Fanuc KAREL source: KT00616.KL

PROGRAM KT00616
%NOLOCKGROUP
VAR
  B1: BOOLEAN
  B2: BOOLEAN
  OUT: INTEGER
BEGIN
  B1 = TRUE
  B2 = FALSE
  B1 = TRUE
  B2 = FALSE
  OUT = NOT B1
END KT00616
